// TIA Portal V21 export
// export: Created 2026-11-11T00:47:52.373981Z, ExportSetting WithDefaults, DisplayName Totally Integrated Automation Portal, DisplayVersion V21 Update 3, DisplayName STEP 7 Professional, DisplayVersion V21 Update 3, DisplayName STEP 7 Safety, DisplayVersion V21, DisplayName Tech WebApplication, DisplayVersion V21, DisplayName WinCC Basic/Comfort/Advanced, DisplayVersion V21 Update 3, DisplayName WinCC Unified, DisplayVersion V21 Update 3
FUNCTION_BLOCK "FB_Lad_TrcvC"   // FB351, LAD
{ S7_Optimized_Access := 'TRUE' }
VERSION : 0.1
// stored: AutoNumber true, IsIECCheckEnabled false, IsRetainMemResEnabled false, MemoryReserve 100, SetENOAutomatically false, UDAEnableTagReadback false
   VAR_INPUT
      en_r : Bool;
      cont : Bool;
      len : UInt;
      id : CONN_OUC;
      adhoc : Bool;
   END_VAR
   VAR_OUTPUT
      done : Bool;
      busy : Bool;
      err : Bool;
      status : Word;
      rcvdlen : UInt;
   END_VAR
   VAR_IN_OUT
      connect : TCON_IP_v4;
      data : Array[0..99] of Byte;
      comrst : Bool;
      addr : Variant;
   END_VAR
   VAR
      inst { S7_SetPoint := 'True'} : TRCV_C;
   END_VAR
BEGIN

REGION Network 1: TRCV_C
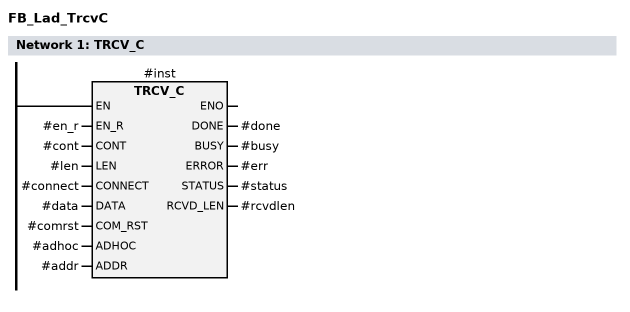
   RUNG wire#powerrail
      #inst.TRCV_C(EN_R := #en_r, CONT := #cont, LEN := #len, CONNECT := #connect, DATA := #data, COM_RST := #comrst, DONE => #done, BUSY => #busy, ERROR => #err, STATUS => #status, RCVD_LEN => #rcvdlen, ADHOC := #adhoc, ADDR := #addr)
   END_RUNG
   // the same network as SCL:
   #inst(EN_R := #en_r,   // TRCV_C
         CONT := #cont,
         LEN := #len,
         CONNECT := #connect,
         DATA := #data,
         COM_RST := #comrst,
         ADHOC := #adhoc,
         ADDR := #addr,
         DONE => #done,
         BUSY => #busy,
         ERROR => #err,
         STATUS => #status,
         RCVD_LEN => #rcvdlen);
END_REGION
END_FUNCTION_BLOCK
